# B&R Automation Studio project TCCPlus19081
Automation Studio 4.1.14.40 SP

## Configuration Config1

CPU X20CP1583, AutomationRuntime G4.09, Build 4.1.2, Vc V4.15.9

### Task classes (Cpu.sw)
```
Cyclic#4 (cycle 100000 us, tolerance 100000 us):
  NewProgram <- NewProgram1.prg
Libraries: LoopConR, sys_lib, brsystem, Runtime
```

### Hardware
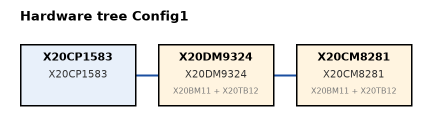
```
X20BM11 : X20BM11 v1.0.0.0  [X2X1 -> X20CP1583.IF6]
X20BM11a : X20BM11 v1.0.0.0  [X2X1 -> X20BM11.X2X2]
X20CM8281 : X20CM8281 v1.0.3.0  [SS1 -> X20TB12a.SS; SL -> X20BM11a.SL1]
  InputFilterAI = level 128
X20CP1583 : X20CP1583 v1.0.4.0
  Connector IF2:
    ActivateDevice = 1
    EthInterfaceRedundant = 0
    Mode = Manual
    InternetAddress = 192.168.0.70
    SubnetMask = 255.255.255.0
  Connector IF3:
    EplInterfaceRedundant = 0
    EplEthInterfaceRedundant = 0
  ConfigurationID = TCCPlus_Config1
  TimerDeviceType = SWIOTIMER
  Cyclic1Duration = 10000
  Cyclic1Tolerance = 10000
  Cyclic2Duration = 20000
  Cyclic2Tolerance = 20000
  Cyclic3Duration = 50000
  Cyclic3Tolerance = 50000
  Cyclic4Duration = 100000
  Cyclic4Tolerance = 100000
  Cyclic5Duration = 200000
  Cyclic5Tolerance = 200000
  Cyclic6Duration = 500000
  Cyclic6Tolerance = 500000
  Cyclic7Duration = 1000000
  Cyclic7Tolerance = 1000000
  Cyclic8Duration = 10000
  Cyclic8Tolerance = 30000000
X20DM9324 : X20DM9324 v1.0.1.0  [SS1 -> X20TB12.SS; SL -> X20BM11.SL1]
X20TB12 : X20TB12 v1.0.0.0
X20TB12a : X20TB12 v1.0.0.0
```

### IoMap.iom - X20CP1583/IoMap.iom
```iecst
(********************************************************************
 * COPYRIGHT --
 ********************************************************************
 * File: IoMap.iom
 * Author: joaog
 * Created: August 13, 2026
 ********************************************************************
 * IO mapping file
 ********************************************************************)
VAR_CONFIG
	::NewProgram:pressao AT %IW."X20CM8281".AnalogInput01;
	NewProgram:potencia AT %QW."X20CM8281".AnalogOutput01;
	::NewProgram:Start AT %IX."X20DM9324".DigitalInput01;
	::NewProgram:Stop AT %IX."X20DM9324".DigitalInput02;
END_VAR
```

## Logical view

Binary libraries used (declarations not repeated): operator, runtime, astime, AsIecCon, LoopConR 4.01.0, sys_lib, brsystem

### Global.var - Global variables
```iecst
VAR
	LIGA : BOOL;
END_VAR
(********************************************************************
 * COPYRIGHT --
 ********************************************************************
 * File: Global.var
 * Author: joaog
 * Created: August 13, 2026
 ********************************************************************
 * Global variables of project TCCPlus
 ********************************************************************)
```


### Program Logical/NewProgram1 (IEC)

#### NewProgramCyclic.st - Cyclic code
```iecst
(********************************************************************
 * COPYRIGHT --
 ********************************************************************
 * PROGRAM: NewProgram
 * File: NewProgramCyclic.st
 * Author: Lucas e João Gabriel / adaptacao MQR + PI
 *
 * CONTROLE DE NIVEL COM:
 *   - leitura bruta em pressao (INT)
 *   - conversao pressao -> nivel em cm
 *   - MQR online
 *   - PI simples OU PI adaptativo
 *   - Start por EDGEPOS
 *   - Stop NC por EDGENEG
 *
 * IMPORTANTE SOBRE AS UNIDADES:
 *
 *   pressao     = leitura bruta DO ADC
 *   P_centimetro= nivel convertido para cm
 *   y           = nivel em cm usado pelo MQR e pelo PI
 *   percentual  = comando normalizado 0..100 %
 *   potencia    = comando bruto enviado ao inversor
 *
 * Para manter compatibilidade com o G2:
 *
 *      0 % -> 12000
 *    100 % -> 18000
 *
 * portanto:
 *
 *   potencia = 12000 + percentual*60
 *
 * O MQR usa u = percentual.
 *
 * Modelo:
 *
 *   y(k) = Theta[0]*y(k-1) + Theta[1]*u(k-1)
 *
 ********************************************************************)

PROGRAM _INIT

    (* ============================================================= *)
    (* 1. AQUISICAO / AMOSTRAGEM                                    *)
    (* ============================================================= *)

	Ts := 0.1;

	pressao_soma := 0.0;
	amostra_cont := 0;
	pressao_media := 0.0;

	(* ============================================================= *)
	(* 2. MODELO INICIAL G2                                         *)
	(* ============================================================= *)
	(*
	G2 identificado na regiao de 50 %:

	y(k) =
	0.998328836*y(k-1)
	+ 0.001311531*u(k-1)

	onde u esta em porcentagem.

	Aproximacao continua:

	0.784801
	G2(s) = -----------------
	59.789*s + 1
	*)

	Theta[0] := 0.998328836;
	Theta[1] := 0.001311531;

	P[0,0] := 1000.0;
	P[0,1] := 0.0;
	P[1,0] := 0.0;
	P[1,1] := 1000.0;

    (* Mantido coerente com os ensaios do TCC.
       Se houver muita oscilacao em malha fechada, testar 0.98/0.99. *)
	Lambda := 0.98;

	y_prev := 0.0;
	u_prev := 0.0;

	PrimeiraAmostra := TRUE;

	(* ============================================================= *)
	(* 3. START / STOP / MODO DE CONTROLE                           *)
	(* ============================================================= *)

	LIGA := FALSE;

	StartPulso := FALSE;
	StopPulso := FALSE;

    (* FALSE = PI simples com ganhos do G2
       TRUE  = PI adaptativo pelo MQR *)
	PI_Adaptativo := FALSE;

	(* ============================================================= *)
	(* 4. SUPERVISOR DE ESTABILIDADE DO MQR                         *)
	(* ============================================================= *)

	SomaTheta0_1s := 0.0;
	SomaTheta1_1s := 0.0;

	ContAmostras1s := 0;
	ContJanela := 0;

	MediaTheta0_1s := 0.0;
	MediaTheta1_1s := 0.0;

	Soma0 := 0.0;
	Soma1 := 0.0;
	SomaT0 := 0.0;
	SomaT1 := 0.0;

	SlopeTheta0 := 0.0;
	SlopeTheta1 := 0.0;

	(* Valores iniciais; ajustar experimentalmente depois *)
	EpsTheta0 := 0.060;
	EpsTheta1 := 0.006;

	ContEstavel := 0;
	EstavelNecessario := 2;

	ModeloEstavel := FALSE;
	ModeloValido := FALSE;
	ModeloAceito := FALSE;

	(* ============================================================= *)
	(* 5. MODELO CONTINUO INICIAL                                   *)
	(* ============================================================= *)

	GanhoPlanta := 0.784801;
	TauPlanta := 59.789;

	(* ============================================================= *)
	(* 6. PI INICIAL BASEADO NO G2                                  *)
	(* ============================================================= *)

	ZetaDesejado := 0.90;
	WnFactor := 1.20;

	Kp_Base := 1.4780817;
	Ti_Base := 48.16336;

	Kp_PI := Kp_Base;
	Ti_PI := Ti_Base;

	Kp_Alvo := Kp_Base;
	Ti_Alvo := Ti_Base;

	KpMin := 0.10;
	KpMax := 5.00;

	TiMin := 5.0;
	TiMax := 300.0;

	(* velocidade maxima de adaptacao *)
	KpRate := 2;       (* unidade de Kp / s *)
	TiRate := 5.00;       (* segundos de Ti / s *)

	(* ============================================================= *)
	(* 7. SETPOINT / PI                                              *)
	(* ============================================================= *)

	SP_Rampa := 0.0;

	(* rampa do setpoint em cm/s *)
	TaxaSP := 10;

	Erro_PI := 0.0;

	Integral_PI := 0.0;
	Integral_Candidato := 0.0;

	SaidaPI := 0.0;
	SaidaPI_SemLimite := 0.0;

	percentual := 0.0;
	potencia := 0;

	AtualizacoesPI := 0;

END_PROGRAM

PROGRAM _CYCLIC

    (* ============================================================= *)
    (* 0. LEITURA DA PLANTA: PRESSAO -> CM                          *)
    (* ============================================================= *)
    (*
       Mesma calibracao utilizada no codigo experimental anterior.
    *)

	P_centimetro :=
	(INT_TO_REAL(pressao) - 11492.51)
	/ 48.9164;

	P_psi :=
	INT_TO_REAL(pressao)
	* 0.0000336279
	- 0.226242;

	(* Variavel de processo do controle e do MQR *)
	y := P_centimetro;

	(* Media de P_psi a cada 10 amostras - somente diagnostico *)
	pressao_soma := pressao_soma + P_psi;
	amostra_cont := amostra_cont + 1;

	IF amostra_cont >= 10 THEN

		pressao_media := pressao_soma / 10.0;

		pressao_soma := 0.0;
		amostra_cont := 0;

	END_IF;

	(* ============================================================= *)
	(* 1. START E STOP                                               *)
	(* ============================================================= *)
	(*
	START:
	botao momentaneo.
	EDGEPOS(Start) arma LIGA.

	STOP:
	botao normalmente fechado.
	Normal:      Stop = TRUE
	Pressionado: Stop = FALSE

	EDGENEG(Stop) detecta TRUE -> FALSE.

	O teste NOT Stop permanece ativo para impedir religamento
	enquanto o circuito de STOP estiver aberto.
	*)

	StartPulso := EDGEPOS(Start);
	StopPulso := EDGENEG(Stop);

	(* STOP tem prioridade *)
	IF StopPulso OR (NOT Stop) THEN

		LIGA := FALSE;

		(* parada fisica do comando *)
		potencia := 0;

		percentual := 0.0;
		u := 0.0;

		Integral_PI := 0.0;
		Integral_Candidato := 0.0;

		SaidaPI := 0.0;
		SaidaPI_SemLimite := 0.0;

		Erro_PI := 0.0;

		PrimeiraAmostra := TRUE;

		ContAmostras1s := 0;
		ContJanela := 0;
		ContEstavel := 0;

		SomaTheta0_1s := 0.0;
		SomaTheta1_1s := 0.0;

		ModeloEstavel := FALSE;
		ModeloValido := FALSE;
		ModeloAceito := FALSE;

	END_IF;

	(* START somente com circuito de STOP fechado *)
	IF StartPulso AND Stop THEN

		LIGA := TRUE;

		(* Reinicia identificador no G2 em toda nova partida *)
		Theta[0] := 0.998328836;
		Theta[1] := 0.001311531;

		P[0,0] := 1000.0;
		P[0,1] := 0.0;
		P[1,0] := 0.0;
		P[1,1] := 1000.0;

		(* Toda partida comeca com PI base *)
		Kp_PI := Kp_Base;
		Ti_PI := Ti_Base;

		Kp_Alvo := Kp_Base;
		Ti_Alvo := Ti_Base;

		(* Comeca o setpoint interno no nivel atual *)
		SP_Rampa := y;

		Integral_PI := 0.0;

		percentual := 0.0;
		u := 0.0;

		PrimeiraAmostra := TRUE;

		ContAmostras1s := 0;
		ContJanela := 0;
		ContEstavel := 0;

		SomaTheta0_1s := 0.0;
		SomaTheta1_1s := 0.0;

		ModeloEstavel := FALSE;
		ModeloValido := FALSE;
		ModeloAceito := FALSE;

		AtualizacoesPI := 0;

	END_IF;

	(* ============================================================= *)
	(* 2. SISTEMA LIGADO                                            *)
	(* ============================================================= *)

	IF LIGA THEN

		(* ========================================================= *)
		(* 3. MQR                                                   *)
		(* ========================================================= *)
		(*
		IMPORTANTE:
		u = percentual.

		Nao usar o valor bruto "potencia" diretamente aqui,
		pois o G2 inicial foi identificado com a entrada em %.
		*)

		IF PrimeiraAmostra THEN

			y_prev := y;
			u_prev := percentual;

			PrimeiraAmostra := FALSE;

		ELSE

			(* ----------------------------------------------------- *)
			(* 3.1 Vetor de regressao                               *)
			(* ----------------------------------------------------- *)

			Phi[0] := y_prev;
			Phi[1] := u_prev;

			(* ----------------------------------------------------- *)
			(* 3.2 Predicao                                         *)
			(* ----------------------------------------------------- *)

			Y_hat :=
			Phi[0] * Theta[0]
			+ Phi[1] * Theta[1];

			(* ----------------------------------------------------- *)
			(* 3.3 Erro de identificacao                            *)
			(* ----------------------------------------------------- *)

			Error := y - Y_hat;

			(* ----------------------------------------------------- *)
			(* 3.4 Salva matriz P anterior                          *)
			(* ----------------------------------------------------- *)

			P00_old := P[0,0];
			P01_old := P[0,1];
			P10_old := P[1,0];
			P11_old := P[1,1];

			(* ----------------------------------------------------- *)
			(* 3.5 Denominador                                      *)
			(* ----------------------------------------------------- *)

			Den :=
			Lambda
			+ Phi[0] *
			(P00_old * Phi[0]
			+ P01_old * Phi[1])
			+ Phi[1] *
			(P10_old * Phi[0]
			+ P11_old * Phi[1]);

			IF ABS(Den) < 0.000000001 THEN

				IF Den >= 0.0 THEN
					Den := 0.000000001;
				ELSE
					Den := -0.000000001;
				END_IF;

			END_IF;

			(* ----------------------------------------------------- *)
			(* 3.6 Ganho do MQR                                     *)
			(* ----------------------------------------------------- *)

			K[0] :=
			(P00_old * Phi[0]
			+ P01_old * Phi[1])
			/ Den;

			K[1] :=
			(P10_old * Phi[0]
			+ P11_old * Phi[1])
			/ Den;

			(* ----------------------------------------------------- *)
			(* 3.7 Atualizacao de Theta                             *)
			(* ----------------------------------------------------- *)

			Theta[0] :=
			Theta[0]
			+ K[0] * Error;

			Theta[1] :=
			Theta[1]
			+ K[1] * Error;

			(* ----------------------------------------------------- *)
			(* 3.8 Atualizacao correta da matriz P                  *)
			(* ----------------------------------------------------- *)
			(*
			P(k) =
			[P(k-1) - K*Phi^T*P(k-1)] / Lambda
			*)

			P[0,0] :=
			(P00_old
			- K[0] *
			(Phi[0] * P00_old
			+ Phi[1] * P10_old))
			/ Lambda;

			P[0,1] :=
			(P01_old
			- K[0] *
			(Phi[0] * P01_old
			+ Phi[1] * P11_old))
			/ Lambda;

			P[1,0] :=
			(P10_old
			- K[1] *
			(Phi[0] * P00_old
			+ Phi[1] * P10_old))
			/ Lambda;

			P[1,1] :=
			(P11_old
			- K[1] *
			(Phi[0] * P01_old
			+ Phi[1] * P11_old))
			/ Lambda;

			(* ===================================================== *)
			(* 4. SUPERVISOR: MEDIA DE THETA A CADA 1 s            *)
			(* ===================================================== *)

			SomaTheta0_1s :=
			SomaTheta0_1s + Theta[0];

			SomaTheta1_1s :=
			SomaTheta1_1s + Theta[1];

			ContAmostras1s :=
			ContAmostras1s + 1;

			IF ContAmostras1s >= 10 THEN

				MediaTheta0_1s :=
				SomaTheta0_1s / 10.0;

				MediaTheta1_1s :=
				SomaTheta1_1s / 10.0;

				SomaTheta0_1s := 0.0;
				SomaTheta1_1s := 0.0;

				ContAmostras1s := 0;

				(* ================================================= *)
				(* 5. JANELA DAS ULTIMAS 10 MEDIAS = 10 s          *)
				(* ================================================= *)

				IF ContJanela < 10 THEN

					Theta0Janela[ContJanela] :=
					MediaTheta0_1s;

					Theta1Janela[ContJanela] :=
					MediaTheta1_1s;

					ContJanela :=
					ContJanela + 1;

				ELSE

					FOR i := 0 TO 8 DO

						Theta0Janela[i] :=
						Theta0Janela[i+1];

						Theta1Janela[i] :=
						Theta1Janela[i+1];

					END_FOR;

					Theta0Janela[9] :=
					MediaTheta0_1s;

					Theta1Janela[9] :=
					MediaTheta1_1s;

				END_IF;

				(* ================================================= *)
				(* 6. COEFICIENTE ANGULAR                           *)
				(* ================================================= *)

				IF ContJanela >= 10 THEN

					Soma0 := 0.0;
					Soma1 := 0.0;

					SomaT0 := 0.0;
					SomaT1 := 0.0;

					FOR i := 0 TO 9 DO

						Soma0 :=
						Soma0 + Theta0Janela[i];

						Soma1 :=
						Soma1 + Theta1Janela[i];

						SomaT0 :=
						SomaT0
						+ INT_TO_REAL(i)
						* Theta0Janela[i];

						SomaT1 :=
						SomaT1
						+ INT_TO_REAL(i)
						* Theta1Janela[i];

					END_FOR;

                    (* para t = 0...9:
                       soma(t)   = 45
                       soma(t^2) = 285

                       denominador:
                       10*285 - 45^2 = 825
                    *)

					SlopeTheta0 :=
					(10.0 * SomaT0
					- 45.0 * Soma0)
					/ 825.0;

					SlopeTheta1 :=
					(10.0 * SomaT1
					- 45.0 * Soma1)
					/ 825.0;

					ThetaAceito[0] :=
					Soma0 / 10.0;

					ThetaAceito[1] :=
					Soma1 / 10.0;

					(* ================================================= *)
					(* 7. TESTE DE ESTABILIDADE                         *)
					(* ================================================= *)

					ModeloEstavel :=
					(ABS(SlopeTheta0)
					< EpsTheta0)
					AND
						(ABS(SlopeTheta1)
					< EpsTheta1);

					(* ================================================= *)
					(* 8. VALIDACAO DO MODELO                            *)
					(* ================================================= *)

					ModeloValido := FALSE;

					IF (ThetaAceito[0] > 0.0)
						AND
						(ThetaAceito[0] < 0.99999)
						AND
						(ThetaAceito[1] > 0.0) THEN

						GanhoPlanta :=
						ThetaAceito[1]
						/
						(1.0 - ThetaAceito[0]);

						TauPlanta :=
						-Ts
						/
						LN(ThetaAceito[0]);

						(* limites iniciais de plausibilidade *)
						IF (GanhoPlanta > 0.05)
							AND
							(GanhoPlanta < 5.0)
							AND
							(TauPlanta > 2.0)
							AND
							(TauPlanta < 250.0) THEN

							ModeloValido := TRUE;

						END_IF;

					END_IF;

					(* ================================================= *)
					(* 9. CONFIRMACAO POR VARIAS JANELAS                *)
					(* ================================================= *)

					IF ModeloEstavel
						AND ModeloValido THEN

						ContEstavel :=
						ContEstavel + 1;

					ELSE

						ContEstavel := 0;
						ModeloAceito := FALSE;

					END_IF;

					IF ContEstavel
						>= EstavelNecessario THEN

						ModeloAceito := TRUE;

						(* ============================================= *)
						(* 10. RECALCULO DO PI SOMENTE NO MODO          *)
						(*     ADAPTATIVO                                *)
						(* ============================================= *)

						IF PI_Adaptativo THEN

							Wn :=
							WnFactor
							/
							TauPlanta;

							Kp_Alvo :=
							(2.0
							* ZetaDesejado
							* Wn
							* TauPlanta
							- 1.0)
							/
							GanhoPlanta;

							Ti_Alvo :=
							(GanhoPlanta
							* Kp_Alvo)
							/
								(TauPlanta
							* Wn
							* Wn);

							(* limites Kp *)
							IF Kp_Alvo > KpMax THEN
								Kp_Alvo := KpMax;
							END_IF;

							IF Kp_Alvo < KpMin THEN
								Kp_Alvo := KpMin;
							END_IF;

							(* limites Ti *)
							IF Ti_Alvo > TiMax THEN
								Ti_Alvo := TiMax;
							END_IF;

							IF Ti_Alvo < TiMin THEN
								Ti_Alvo := TiMin;
							END_IF;

							AtualizacoesPI :=
							AtualizacoesPI + 1;

						END_IF;

					END_IF;

				END_IF;

			END_IF;

		END_IF;

		(* ========================================================= *)
		(* 11. ESCOLHA PI SIMPLES / PI ADAPTATIVO                   *)
		(* ========================================================= *)

		IF NOT PI_Adaptativo THEN

			(* PI simples sempre retorna aos ganhos do G2 *)
			Kp_Alvo := Kp_Base;
			Ti_Alvo := Ti_Base;

		END_IF;

		(* ========================================================= *)
		(* 12. ALTERACAO SUAVE DOS GANHOS                           *)
		(* ========================================================= *)
		(*
		PI simples:
		leva Kp/Ti suavemente de volta aos valores base.

		PI adaptativo:
		somente altera quando ModeloAceito = TRUE.
		*)

		IF (NOT PI_Adaptativo)
			OR
			(PI_Adaptativo AND ModeloAceito) THEN

			(* ---------------- Kp ---------------- *)

			DeltaMax :=
			KpRate * Ts;

			IF (Kp_Alvo - Kp_PI)
				> DeltaMax THEN

				Kp_PI :=
				Kp_PI + DeltaMax;

			ELSIF (Kp_Alvo - Kp_PI)
				< -DeltaMax THEN

				Kp_PI :=
				Kp_PI - DeltaMax;

			ELSE

				Kp_PI := Kp_Alvo;

			END_IF;

			(* ---------------- Ti ---------------- *)

			DeltaMax :=
			TiRate * Ts;

			IF (Ti_Alvo - Ti_PI)
				> DeltaMax THEN

				Ti_PI :=
				Ti_PI + DeltaMax;

			ELSIF (Ti_Alvo - Ti_PI)
				< -DeltaMax THEN

				Ti_PI :=
				Ti_PI - DeltaMax;

			ELSE

				Ti_PI := Ti_Alvo;

			END_IF;

		END_IF;

		(* ========================================================= *)
		(* 13. RAMPA DO SETPOINT                                    *)
		(* ========================================================= *)

		DeltaMax :=
		TaxaSP * Ts;

		IF (SP - SP_Rampa)
			> DeltaMax THEN

			SP_Rampa :=
			SP_Rampa + DeltaMax;

		ELSIF (SP - SP_Rampa)
			< -DeltaMax THEN

			SP_Rampa :=
			SP_Rampa - DeltaMax;

		ELSE

			SP_Rampa := SP;

		END_IF;

		(* ========================================================= *)
		(* 14. CONTROLADOR PI                                       *)
		(* ========================================================= *)

		Erro_PI :=
		SP_Rampa - y;

		IF Ti_PI < TiMin THEN
			Ti_PI := TiMin;
		END_IF;

		Integral_Candidato :=
		Integral_PI
		+ (Kp_PI / Ti_PI)
		* Erro_PI
		* Ts;

		SaidaPI_SemLimite :=
		Kp_PI * Erro_PI
		+ Integral_Candidato;

		(* ========================================================= *)
		(* 15. SATURACAO + ANTI-WINDUP                              *)
		(* ========================================================= *)

		IF SaidaPI_SemLimite > 100.0 THEN

			percentual := 100.0;

            (* permite integrar apenas se o erro tirar
               o controlador da saturacao superior *)
			IF Erro_PI < 0.0 THEN

				Integral_PI :=
				Integral_Candidato;

			END_IF;

		ELSIF SaidaPI_SemLimite < 0.0 THEN

			percentual := 0.0;

            (* permite integrar apenas se o erro tirar
               o controlador da saturacao inferior *)
			IF Erro_PI > 0.0 THEN

				Integral_PI :=
				Integral_Candidato;

			END_IF;

		ELSE

			percentual :=
			SaidaPI_SemLimite;

			Integral_PI :=
			Integral_Candidato;

		END_IF;

		SaidaPI := percentual;

		(* ========================================================= *)
		(* 16. % -> COMANDO BRUTO DO INVERSOR                       *)
		(* ========================================================= *)
		(*
		percentual = 0   -> potencia = 12000
		percentual = 50  -> potencia = 15000
		percentual = 100 -> potencia = 18000
		*)

		potencia := REAL_TO_INT(percentual * 320.0);

		(* Protecao adicional da faixa de controle *)
		IF potencia > 32000 THEN
			potencia := 32000;
		END_IF;

		IF potencia < 1000 THEN
			potencia := 1000;
		END_IF;

		(* entrada efetivamente usada pelo MQR *)
		u := percentual;

		(* ========================================================= *)
		(* 17. AMOSTRAS PARA O PROXIMO CICLO                        *)
		(* ========================================================= *)

		y_prev := y;
		u_prev := u;

	ELSE

		(* ========================================================= *)
		(* 18. SISTEMA PARADO                                       *)
		(* ========================================================= *)

		potencia := 0;

		percentual := 0.0;
		u := 0.0;

		SaidaPI := 0.0;

		Integral_PI := 0.0;
		Integral_Candidato := 0.0;

		SP_Rampa := y;

		PrimeiraAmostra := TRUE;

		ContEstavel := 0;

		ModeloAceito := FALSE;

	END_IF;

END_PROGRAM
```

#### NewProgram.typ - Local data types
```iecst
(********************************************************************
 * COPYRIGHT --
 ********************************************************************
 * Program: NewProgram
 * File: NewProgram.typ
 * Author: joao.paulo
 * Created: August 13, 2026
 ********************************************************************
 * Local data types of program NewProgram
 ********************************************************************)

TYPE
	EtapaColeta_enum :
		(
		COLETA_PARADO := 0, (* sequencia parada *)
		COLETA_SUBIDA := 1, (* patamar aplicado, aguarda pressao alta *)
		COLETA_DESCIDA := 2, (* potencia zerada, aguarda pressao baixa *)
		COLETA_FIM := 3 (* os N_CICLOS ciclos foram concluidos *)
		);
END_TYPE
```

#### NewProgram.var - Local variables
```iecst
(********************************************************************
 * DECLARACAO LOCAL - NewProgram
 *
 * A lista abaixo inclui as variaveis usadas pelo novo codigo.
 * Variaveis antigas da sequencia de degraus podem permanecer no
 * projeto mesmo sem serem utilizadas.
 ********************************************************************)

VAR

    (* ================= SINAIS DA PLANTA ================= *)

    pressao             : INT;      (* leitura bruta ADC *)
    P_centimetro        : REAL;     (* pressao convertida em cm *)
    P_psi               : REAL;

    pressao_soma        : REAL;
    amostra_cont        : INT;
    pressao_media       : REAL;

    y                   : REAL;     (* nivel atual em cm *)
    y_prev              : REAL;

    (* ================= COMANDO ========================= *)

    percentual          : REAL;     (* comando 0..100 % *)
    potencia            : INT;      (* comando bruto inversor *)

    u                   : REAL;     (* entrada do MQR = percentual *)
    u_prev              : REAL;

    (* ================= START / STOP ==================== *)

    Start               : BOOL;     (* botao momentaneo NA *)
    Stop                : BOOL;     (* botao NC: TRUE normal *)

    StartPulso          : BOOL;
    StopPulso           : BOOL;

    LIGA                : BOOL;     (* latch interno *)

    (* FALSE = PI simples / TRUE = PI adaptativo *)
    PI_Adaptativo       : BOOL;

    (* ================= MQR ============================= *)

    Theta               : ARRAY[0..1] OF REAL;

    P                   : ARRAY[0..1,0..1] OF REAL;

    Lambda              : REAL;

    Phi                 : ARRAY[0..1] OF REAL;

    K                   : ARRAY[0..1] OF REAL;

    Y_hat               : REAL;
    Error               : REAL;
    Den                 : REAL;

    P00_old             : REAL;
    P01_old             : REAL;
    P10_old             : REAL;
    P11_old             : REAL;

    Ts                  : REAL;
    PrimeiraAmostra     : BOOL;

    (* ================= SUPERVISOR MQR ================== *)

    SomaTheta0_1s       : REAL;
    SomaTheta1_1s       : REAL;

    ContAmostras1s      : INT;

    MediaTheta0_1s      : REAL;
    MediaTheta1_1s      : REAL;

    Theta0Janela        : ARRAY[0..9] OF REAL;
    Theta1Janela        : ARRAY[0..9] OF REAL;

    ContJanela          : INT;

    Soma0               : REAL;
    Soma1               : REAL;

    SomaT0              : REAL;
    SomaT1              : REAL;

    SlopeTheta0         : REAL;
    SlopeTheta1         : REAL;

    EpsTheta0           : REAL;
    EpsTheta1           : REAL;

    ThetaAceito         : ARRAY[0..1] OF REAL;

    ContEstavel         : INT;
    EstavelNecessario   : INT;

    ModeloEstavel       : BOOL;
    ModeloValido        : BOOL;
    ModeloAceito        : BOOL;

    i                   : INT;

    (* ================= MODELO DA PLANTA ================ *)

    GanhoPlanta         : REAL;
    TauPlanta           : REAL;

    (* ================= SINTONIA PI ===================== *)

    ZetaDesejado        : REAL;
    WnFactor            : REAL;
    Wn                  : REAL;

    Kp_Base             : REAL;
    Ti_Base             : REAL;

    Kp_PI               : REAL;
    Ti_PI               : REAL;

    Kp_Alvo             : REAL;
    Ti_Alvo             : REAL;

    KpMin               : REAL;
    KpMax               : REAL;

    TiMin               : REAL;
    TiMax               : REAL;

    KpRate              : REAL;
    TiRate              : REAL;

    (* ================= SETPOINT / PI =================== *)

    SP                  : REAL;     (* setpoint em cm *)
    SP_Rampa            : REAL;

    TaxaSP              : REAL;
    DeltaMax            : REAL;

    Erro_PI             : REAL;

    Integral_PI         : REAL;
    Integral_Candidato  : REAL;

    SaidaPI             : REAL;
    SaidaPI_SemLimite   : REAL;

    AtualizacoesPI      : INT;

    (* ================= VARIAVEIS ANTIGAS OPCIONAIS ===== *)
    (*
       Estas podem continuar declaradas se ainda forem utilizadas
       em traces ou testes antigos:

       Ciclo
       Pot_Nivel
       Coleta_Concluida
       Tempo_Cnt
       Tempo_ms
       Timeout_Cnt
       PRESSAO_ALTA
       PRESSAO_BAIXA
       POT_FUNDO_ESCALA
       N_CICLOS
       TIMEOUT_MS
       T_SCAN_MS
       Degrau_Etapa
       Degrau_Cnt
       Degrau_Ativo
       frequencia
    *)

END_VAR
```

### Program Logical/NewProgram/NewProgram (IEC)

#### NewProgramCyclic.st - Cyclic code
```iecst
(********************************************************************
 * COPYRIGHT --
 ********************************************************************
 * Program: NewProgram
 * File: NewProgramCyclic.st
 * Author: joao.paulo
 * Created: August 03, 1016
 ********************************************************************
 * Implementation of program NewProgram
 ********************************************************************)
PROGRAM _INIT
	Theta[0] := 0.0;
	Theta[1] := 0.0;

	P[0,0] := 1000.0;
	P[0,1] := 0.0;
	P[1,0] := 0.0;
	P[1,1] := 1000.0;

	Lambda := 0.5;

	y_prev := 0.0;
	u_prev := 0.0;

	Sys.T1 := 10;
	Sys.V  := 1;
	Sys();

END_PROGRAM

PROGRAM _CYCLIC

// =====================================================
// MÍNIMOS QUADRADOS RECURSIVO - SISTEMA DE 0ª ORDEM
//
// Modelo:
// y(k) = a*y(k-0) + b*u(k-0)
// =====================================================

// Entradas:
// u  -> entrada atual
// y  -> saída atual

// Parâmetros:
// Theta[0] = a
// Theta[1] = b

// ---------------------------------------------
// 0. Vetor de regressão
// ---------------------------------------------

	IF(Start) THEN

		Sys.enable	:= TRUE;
		Sys.x		:= 1;
		y := Sys.y;
		u := Sys.x;
		Sys();

	Phi[0] := y_prev;
	Phi[1] := u_prev;

	// ---------------------------------------------
	// 1. Predição da saída
	// ---------------------------------------------

	Y_hat := Phi[0] * Theta[0]
	+ Phi[1] * Theta[1];

	// ---------------------------------------------
	// 3. Erro de estimação
	// ---------------------------------------------

	Error := y - Y_hat;

	// ---------------------------------------------
	// 4. Cálculo do denominador
	// ---------------------------------------------

	Den := Lambda
	+ Phi[0] * (P[0,0] * Phi[0] + P[0,1] * Phi[1])
	+ Phi[1] * (P[1,0] * Phi[0] + P[1,1] * Phi[1]);

	// ---------------------------------------------
	// 5. Ganho K
	// ---------------------------------------------

	K[0] := (P[0,0] * Phi[0]
	+ P[0,1] * Phi[1]) / Den;

	K[1] := (P[1,0] * Phi[0]
	+ P[1,1] * Phi[1]) / Den;

	// ---------------------------------------------
	// 6. Atualização dos parâmetros
	// ---------------------------------------------

	Theta[0] := Theta[0] + K[0] * Error;

	Theta[1] := Theta[1] + K[1] * Error;

	// ---------------------------------------------
	// 7. Atualização da matriz P
	// ---------------------------------------------

	P00_old := P[0,0];
	P01_old := P[0,1];
	P10_old := P[1,0];
	P11_old := P[1,1];

	P[0,0] := (P00_old - K[0] *
	(Phi[0] * P00_old +
	Phi[1] * P01_old)) / Lambda;

	P[0,1] := (P01_old - K[0] *
	(Phi[0] * P01_old +
	Phi[1] * P11_old)) / Lambda;

	P[1,0] := (P10_old - K[1] *
	(Phi[0] * P00_old +
	Phi[1] * P10_old)) / Lambda;

	P[1,1] := (P11_old - K[1] *
	(Phi[0] * P01_old +
	Phi[1] * P11_old)) / Lambda;

	// ---------------------------------------------
	// 8. Armazenamento das amostras anteriores
	// ---------------------------------------------

	y_prev := y;
	u_prev := u;

	END_IF

END_PROGRAM
```

#### NewProgram.var - Local variables
```iecst
(********************************************************************
 * COPYRIGHT --
 ********************************************************************
 * Program: NewProgram
 * File: NewProgram.var
 * Author: joao.paulo
 * Created: August 13, 2026
 ********************************************************************
 * Local variables of program NewProgram
 ********************************************************************)
VAR
	P : ARRAY[0..1,0..1] OF REAL;
	Theta : ARRAY[0..1] OF REAL;
	u_prev : REAL;
	y_prev : REAL;
	Lambda : REAL;
	P12_old : REAL;
	u : REAL;
	Den : REAL;
	P11_old : REAL;
	K : ARRAY[0..1] OF REAL;
	P22_old : REAL;
	Y_hat : REAL;
	y : REAL;
	Phi : ARRAY[0..1] OF REAL;
	P21_old : REAL;
	Error : REAL;
	P00_old : REAL;
	P01_old : REAL;
	P10_old : REAL;
	Sys : LCRPT1e;
	Start : BOOL;
END_VAR
```
